// TIA Portal V20 export
// export: Created 2026-10-20T12:39:45.8971226Z, ExportSetting WithDefaults, DisplayName Totally Integrated Automation Portal, DisplayVersion V20 Update 6, DisplayName TIA Portal Openness, DisplayVersion V20 Update 6, DisplayName TIA Portal Version Control Interface, DisplayVersion V20 Update 6, DisplayName SINAMICS Startdrive Advanced, DisplayVersion V20 SP1, DisplayName SINAMICS Startdrive G130, G150, S120, S150, SINAMICS MV, G220, S200, S210, DisplayVersion V20 SP1, DisplayName SINAMICS Startdrive G110M, G120, G120C, G120D, G120P, G115D, DisplayVersion V20 SP1, DisplayName STEP 7 Professional, DisplayVersion V20 Update 6, DisplayName STEP 7 Safety, DisplayVersion V20 Update 2, DisplayName WinCC Basic/Comfort/Advanced, DisplayVersion V20 Update 6, DisplayName WinCC Unified, DisplayVersion V20 Update 6
FUNCTION_BLOCK "Main_Safety_RTG1"   // FB123, F_FBD
{ S7_Optimized_Access := 'TRUE' }
VERSION : 0.1
// stored: AutoNumber false, IsIECCheckEnabled false, UDAEnableTagReadback false
   VAR
      Safety_OK : Bool;
      ACK : Bool;
   END_VAR
   VAR_TEMP
      HMI_1_Estop_Pressed_1 : Bool;
      HMI_1_Estop_Pressed_2 : Bool;
      HMI_1_Estop_Pressed_3 : Bool;
      HMI_1_Estop_Pressed_4 : Bool;
      HMI_1_Estop_Pressed_5 : Bool;
      HMI_2_Estop_Pressed_1 : Bool;
      HMI_2_Estop_Pressed_2 : Bool;
      HMI_2_Estop_Pressed_3 : Bool;
      HMI_2_Estop_Pressed_4 : Bool;
      HMI_2_Estop_Pressed_5 : Bool;
      HMI_1_Reset_Comiss_1 : Bool;
      HMI_1_Reset_Comiss_2 : Bool;
      HMI_1_Reset_Comiss_3 : Bool;
      HMI_1_Reset_Comiss_4 : Bool;
      HMI_1_Reset_Comiss_5 : Bool;
      HMI_2_Reset_Comiss_1 : Bool;
      HMI_2_Reset_Comiss_2 : Bool;
      HMI_2_Reset_Comiss_3 : Bool;
      HMI_2_Reset_Comiss_4 : Bool;
      HMI_2_Reset_Comiss_5 : Bool;
   END_VAR
BEGIN

REGION Network 1: MAIN PANEL
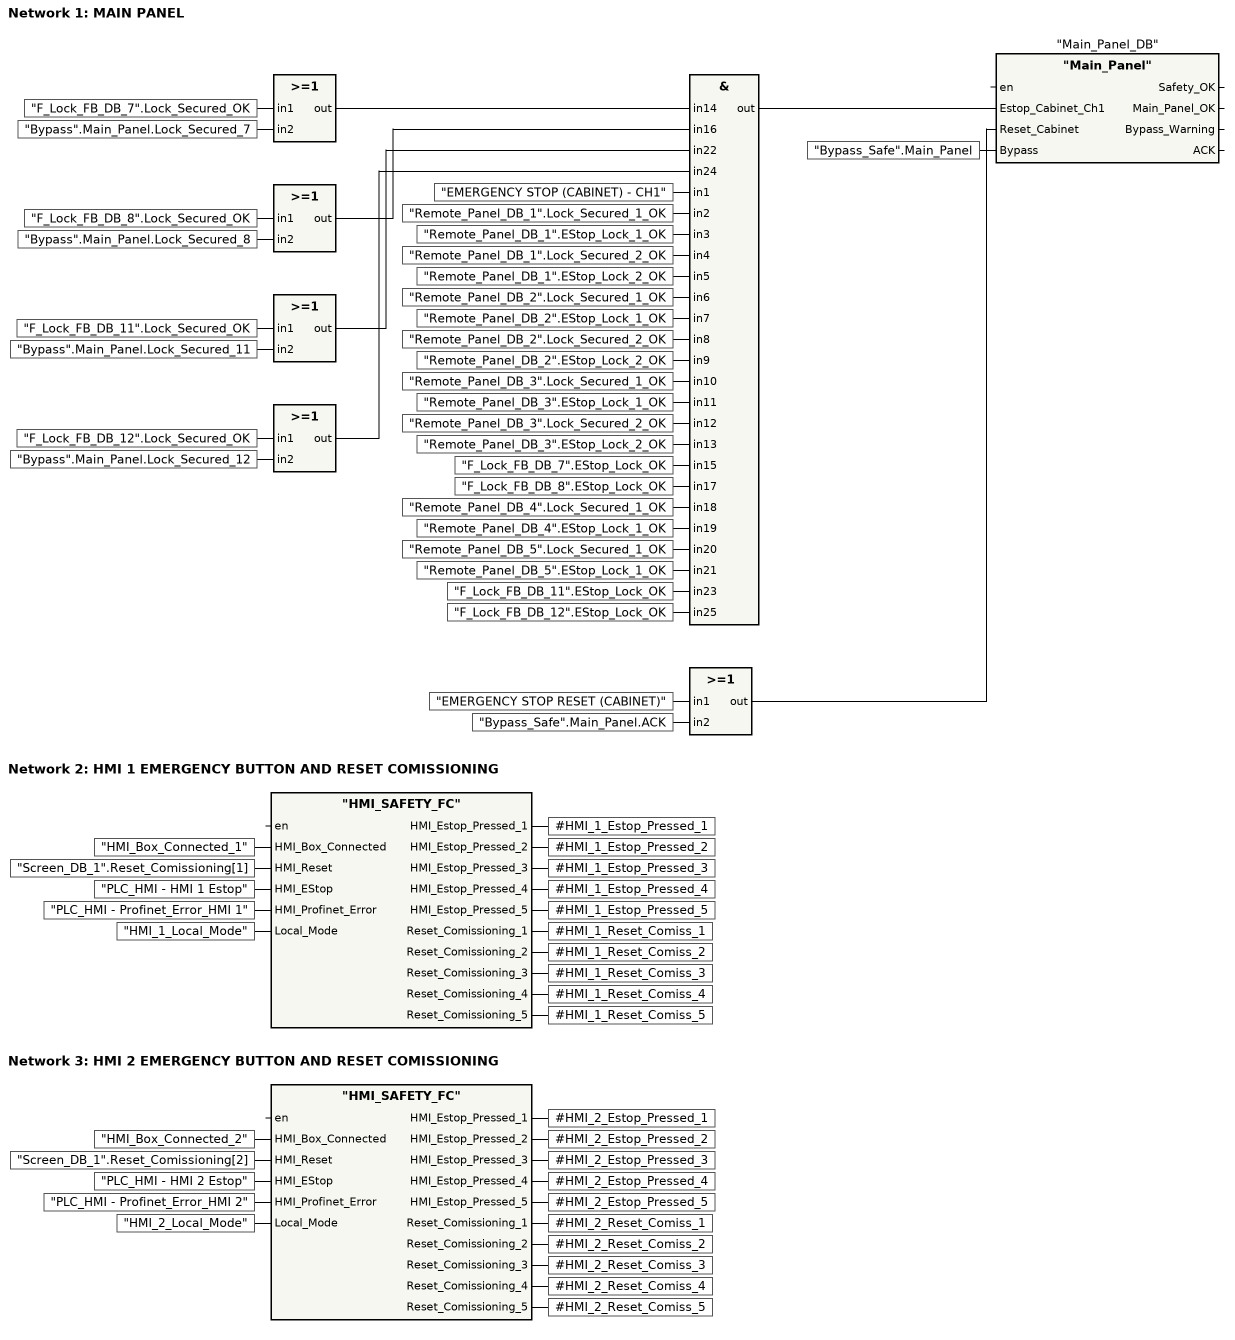
   "Main_Panel_DB"(Estop_Cabinet_Ch1 := ("F_Lock_FB_DB_7".Lock_Secured_OK OR "Bypass".Main_Panel.Lock_Secured_7) AND ("F_Lock_FB_DB_8".Lock_Secured_OK OR "Bypass".Main_Panel.Lock_Secured_8) AND ("F_Lock_FB_DB_11".Lock_Secured_OK OR "Bypass".Main_Panel.Lock_Secured_11) AND ("F_Lock_FB_DB_12".Lock_Secured_OK OR "Bypass".Main_Panel.Lock_Secured_12) AND "EMERGENCY STOP (CABINET) - CH1" AND "Remote_Panel_DB_1".Lock_Secured_1_OK AND "Remote_Panel_DB_1".EStop_Lock_1_OK AND "Remote_Panel_DB_1".Lock_Secured_2_OK AND "Remote_Panel_DB_1".EStop_Lock_2_OK AND "Remote_Panel_DB_2".Lock_Secured_1_OK AND "Remote_Panel_DB_2".EStop_Lock_1_OK AND "Remote_Panel_DB_2".Lock_Secured_2_OK AND "Remote_Panel_DB_2".EStop_Lock_2_OK AND "Remote_Panel_DB_3".Lock_Secured_1_OK AND "Remote_Panel_DB_3".EStop_Lock_1_OK AND "Remote_Panel_DB_3".Lock_Secured_2_OK AND "Remote_Panel_DB_3".EStop_Lock_2_OK AND "F_Lock_FB_DB_7".EStop_Lock_OK AND "F_Lock_FB_DB_8".EStop_Lock_OK AND "Remote_Panel_DB_4".Lock_Secured_1_OK AND "Remote_Panel_DB_4".EStop_Lock_1_OK AND "Remote_Panel_DB_5".Lock_Secured_1_OK AND "Remote_Panel_DB_5".EStop_Lock_1_OK AND "F_Lock_FB_DB_11".EStop_Lock_OK AND "F_Lock_FB_DB_12".EStop_Lock_OK,   // "Main_Panel"
                   Reset_Cabinet := "EMERGENCY STOP RESET (CABINET)" OR "Bypass_Safe".Main_Panel.ACK,
                   Bypass := "Bypass_Safe".Main_Panel);
END_REGION

REGION Network 2: HMI 1 EMERGENCY BUTTON AND RESET COMISSIONING
   "HMI_SAFETY_FC"(HMI_Box_Connected := "HMI_Box_Connected_1",
                   HMI_Reset := "Screen_DB_1".Reset_Comissioning[1],
                   HMI_EStop := "PLC_HMI - HMI 1 Estop",
                   HMI_Profinet_Error := "PLC_HMI - Profinet_Error_HMI 1",
                   Local_Mode := "HMI_1_Local_Mode",
                   HMI_Estop_Pressed_1 => #HMI_1_Estop_Pressed_1,
                   HMI_Estop_Pressed_2 => #HMI_1_Estop_Pressed_2,
                   HMI_Estop_Pressed_3 => #HMI_1_Estop_Pressed_3,
                   HMI_Estop_Pressed_4 => #HMI_1_Estop_Pressed_4,
                   HMI_Estop_Pressed_5 => #HMI_1_Estop_Pressed_5,
                   Reset_Comissioning_1 => #HMI_1_Reset_Comiss_1,
                   Reset_Comissioning_2 => #HMI_1_Reset_Comiss_2,
                   Reset_Comissioning_3 => #HMI_1_Reset_Comiss_3,
                   Reset_Comissioning_4 => #HMI_1_Reset_Comiss_4,
                   Reset_Comissioning_5 => #HMI_1_Reset_Comiss_5);
END_REGION

REGION Network 3: HMI 2 EMERGENCY BUTTON AND RESET COMISSIONING
   "HMI_SAFETY_FC"(HMI_Box_Connected := "HMI_Box_Connected_2",
                   HMI_Reset := "Screen_DB_1".Reset_Comissioning[2],
                   HMI_EStop := "PLC_HMI - HMI 2 Estop",
                   HMI_Profinet_Error := "PLC_HMI - Profinet_Error_HMI 2",
                   Local_Mode := "HMI_2_Local_Mode",
                   HMI_Estop_Pressed_1 => #HMI_2_Estop_Pressed_1,
                   HMI_Estop_Pressed_2 => #HMI_2_Estop_Pressed_2,
                   HMI_Estop_Pressed_3 => #HMI_2_Estop_Pressed_3,
                   HMI_Estop_Pressed_4 => #HMI_2_Estop_Pressed_4,
                   HMI_Estop_Pressed_5 => #HMI_2_Estop_Pressed_5,
                   Reset_Comissioning_1 => #HMI_2_Reset_Comiss_1,
                   Reset_Comissioning_2 => #HMI_2_Reset_Comiss_2,
                   Reset_Comissioning_3 => #HMI_2_Reset_Comiss_3,
                   Reset_Comissioning_4 => #HMI_2_Reset_Comiss_4,
                   Reset_Comissioning_5 => #HMI_2_Reset_Comiss_5);
END_REGION

REGION Network 4: Remote Panel 1
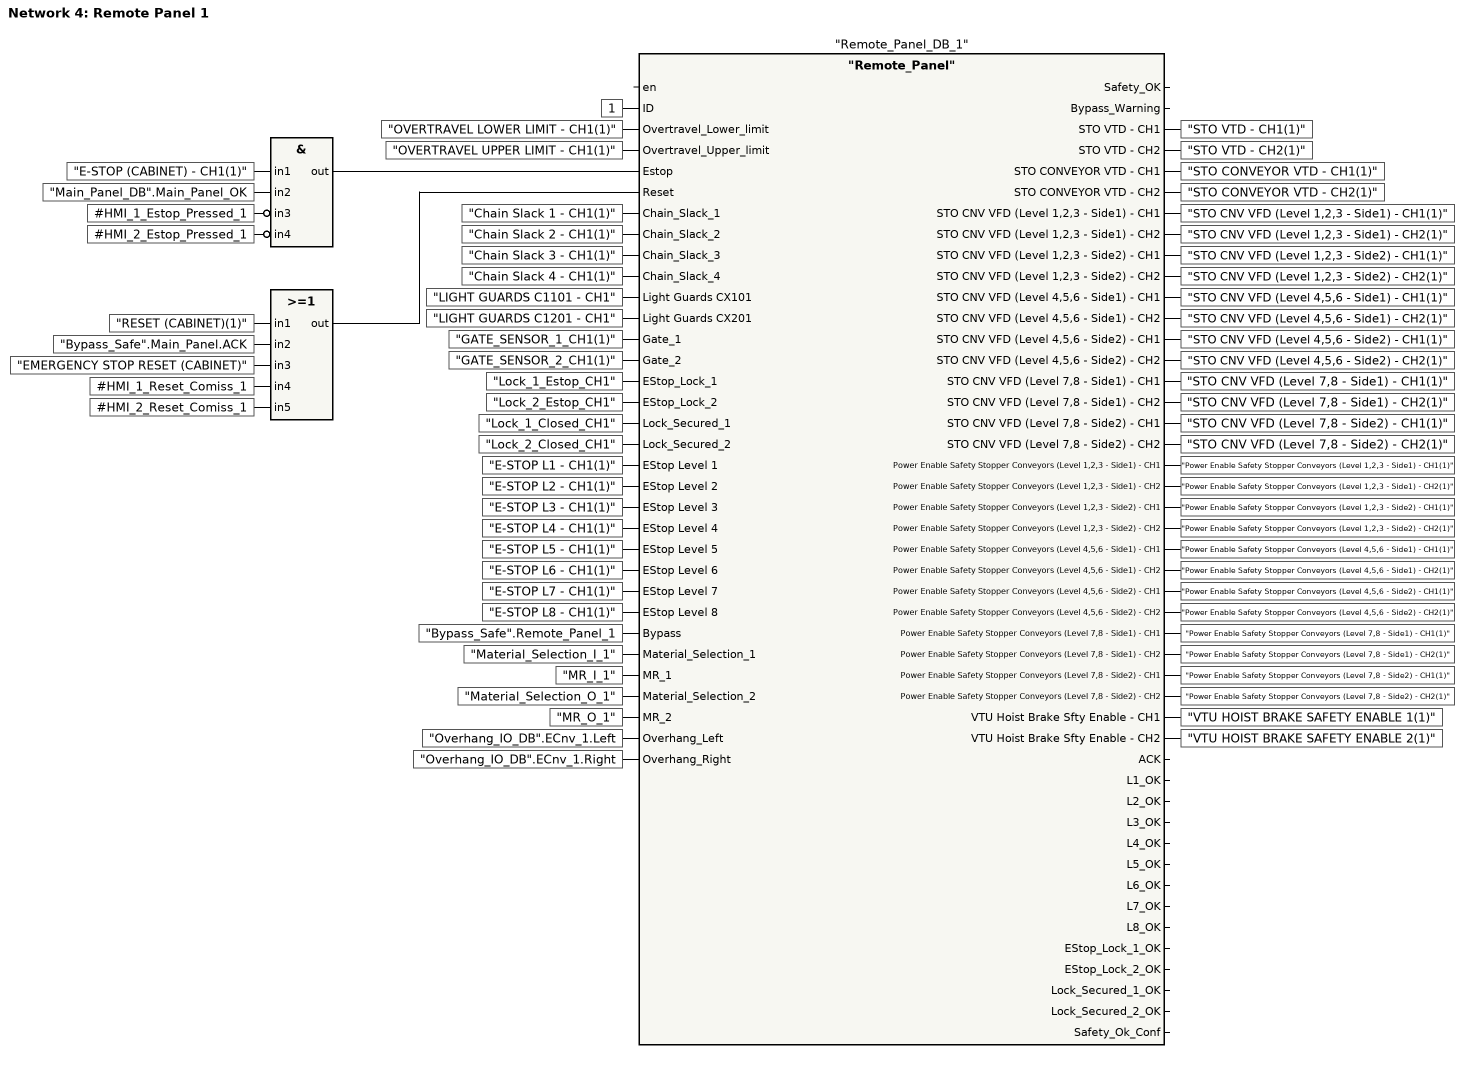
   "Remote_Panel_DB_1"(ID := 1,   // "Remote_Panel"
                       Overtravel_Lower_limit := "OVERTRAVEL LOWER LIMIT - CH1(1)",
                       Overtravel_Upper_limit := "OVERTRAVEL UPPER LIMIT - CH1(1)",
                       Estop := "E-STOP (CABINET) - CH1(1)" AND "Main_Panel_DB".Main_Panel_OK AND NOT #HMI_1_Estop_Pressed_1 AND NOT #HMI_2_Estop_Pressed_1,
                       Reset := "RESET (CABINET)(1)" OR "Bypass_Safe".Main_Panel.ACK OR "EMERGENCY STOP RESET (CABINET)" OR #HMI_1_Reset_Comiss_1 OR #HMI_2_Reset_Comiss_1,
                       Chain_Slack_1 := "Chain Slack 1 - CH1(1)",
                       Chain_Slack_2 := "Chain Slack 2 - CH1(1)",
                       Chain_Slack_3 := "Chain Slack 3 - CH1(1)",
                       Chain_Slack_4 := "Chain Slack 4 - CH1(1)",
                       "Light Guards CX101" := "LIGHT GUARDS C1101 - CH1",
                       "Light Guards CX201" := "LIGHT GUARDS C1201 - CH1",
                       Gate_1 := "GATE_SENSOR_1_CH1(1)",
                       Gate_2 := "GATE_SENSOR_2_CH1(1)",
                       EStop_Lock_1 := "Lock_1_Estop_CH1",
                       EStop_Lock_2 := "Lock_2_Estop_CH1",
                       Lock_Secured_1 := "Lock_1_Closed_CH1",
                       Lock_Secured_2 := "Lock_2_Closed_CH1",
                       "EStop Level 1" := "E-STOP L1 - CH1(1)",
                       "EStop Level 2" := "E-STOP L2 - CH1(1)",
                       "EStop Level 3" := "E-STOP L3 - CH1(1)",
                       "EStop Level 4" := "E-STOP L4 - CH1(1)",
                       "EStop Level 5" := "E-STOP L5 - CH1(1)",
                       "EStop Level 6" := "E-STOP L6 - CH1(1)",
                       "EStop Level 7" := "E-STOP L7 - CH1(1)",
                       "EStop Level 8" := "E-STOP L8 - CH1(1)",
                       Bypass := "Bypass_Safe".Remote_Panel_1,
                       Material_Selection_1 := "Material_Selection_I_1",
                       MR_1 := "MR_I_1",
                       Material_Selection_2 := "Material_Selection_O_1",
                       MR_2 := "MR_O_1",
                       Overhang_Left := "Overhang_IO_DB".ECnv_1.Left,
                       Overhang_Right := "Overhang_IO_DB".ECnv_1.Right,
                       "STO VTD - CH1" => "STO VTD - CH1(1)",
                       "STO VTD - CH2" => "STO VTD - CH2(1)",
                       "STO CONVEYOR VTD - CH1" => "STO CONVEYOR VTD - CH1(1)",
                       "STO CONVEYOR VTD - CH2" => "STO CONVEYOR VTD - CH2(1)",
                       "STO CNV VFD (Level 1,2,3 - Side1) - CH1" => "STO CNV VFD (Level 1,2,3 - Side1) - CH1(1)",
                       "STO CNV VFD (Level 1,2,3 - Side1) - CH2" => "STO CNV VFD (Level 1,2,3 - Side1) - CH2(1)",
                       "STO CNV VFD (Level 1,2,3 - Side2) - CH1" => "STO CNV VFD (Level 1,2,3 - Side2) - CH1(1)",
                       "STO CNV VFD (Level 1,2,3 - Side2) - CH2" => "STO CNV VFD (Level 1,2,3 - Side2) - CH2(1)",
                       "STO CNV VFD (Level 4,5,6 - Side1) - CH1" => "STO CNV VFD (Level 4,5,6 - Side1) - CH1(1)",
                       "STO CNV VFD (Level 4,5,6 - Side1) - CH2" => "STO CNV VFD (Level 4,5,6 - Side1) - CH2(1)",
                       "STO CNV VFD (Level 4,5,6 - Side2) - CH1" => "STO CNV VFD (Level 4,5,6 - Side2) - CH1(1)",
                       "STO CNV VFD (Level 4,5,6 - Side2) - CH2" => "STO CNV VFD (Level 4,5,6 - Side2) - CH2(1)",
                       "STO CNV VFD (Level 7,8 - Side1) - CH1" => "STO CNV VFD (Level 7,8 - Side1) - CH1(1)",
                       "STO CNV VFD (Level 7,8 - Side1) - CH2" => "STO CNV VFD (Level 7,8 - Side1) - CH2(1)",
                       "STO CNV VFD (Level 7,8 - Side2) - CH1" => "STO CNV VFD (Level 7,8 - Side2) - CH1(1)",
                       "STO CNV VFD (Level 7,8 - Side2) - CH2" => "STO CNV VFD (Level 7,8 - Side2) - CH2(1)",
                       "Power Enable Safety Stopper Conveyors (Level 1,2,3 - Side1) - CH1" => "Power Enable Safety Stopper Conveyors (Level 1,2,3 - Side1) - CH1(1)",
                       "Power Enable Safety Stopper Conveyors (Level 1,2,3 - Side1) - CH2" => "Power Enable Safety Stopper Conveyors (Level 1,2,3 - Side1) - CH2(1)",
                       "Power Enable Safety Stopper Conveyors (Level 1,2,3 - Side2) - CH1" => "Power Enable Safety Stopper Conveyors (Level 1,2,3 - Side2) - CH1(1)",
                       "Power Enable Safety Stopper Conveyors (Level 1,2,3 - Side2) - CH2" => "Power Enable Safety Stopper Conveyors (Level 1,2,3 - Side2) - CH2(1)",
                       "Power Enable Safety Stopper Conveyors (Level 4,5,6 - Side1) - CH1" => "Power Enable Safety Stopper Conveyors (Level 4,5,6 - Side1) - CH1(1)",
                       "Power Enable Safety Stopper Conveyors (Level 4,5,6 - Side1) - CH2" => "Power Enable Safety Stopper Conveyors (Level 4,5,6 - Side1) - CH2(1)",
                       "Power Enable Safety Stopper Conveyors (Level 4,5,6 - Side2) - CH1" => "Power Enable Safety Stopper Conveyors (Level 4,5,6 - Side2) - CH1(1)",
                       "Power Enable Safety Stopper Conveyors (Level 4,5,6 - Side2) - CH2" => "Power Enable Safety Stopper Conveyors (Level 4,5,6 - Side2) - CH2(1)",
                       "Power Enable Safety Stopper Conveyors (Level 7,8 - Side1) - CH1" => "Power Enable Safety Stopper Conveyors (Level 7,8 - Side1) - CH1(1)",
                       "Power Enable Safety Stopper Conveyors (Level 7,8 - Side1) - CH2" => "Power Enable Safety Stopper Conveyors (Level 7,8 - Side1) - CH2(1)",
                       "Power Enable Safety Stopper Conveyors (Level 7,8 - Side2) - CH1" => "Power Enable Safety Stopper Conveyors (Level 7,8 - Side2) - CH1(1)",
                       "Power Enable Safety Stopper Conveyors (Level 7,8 - Side2) - CH2" => "Power Enable Safety Stopper Conveyors (Level 7,8 - Side2) - CH2(1)",
                       "VTU Hoist Brake Sfty Enable - CH1" => "VTU HOIST BRAKE SAFETY ENABLE 1(1)",
                       "VTU Hoist Brake Sfty Enable - CH2" => "VTU HOIST BRAKE SAFETY ENABLE 2(1)");
END_REGION

REGION Network 5: Remote Panel 2
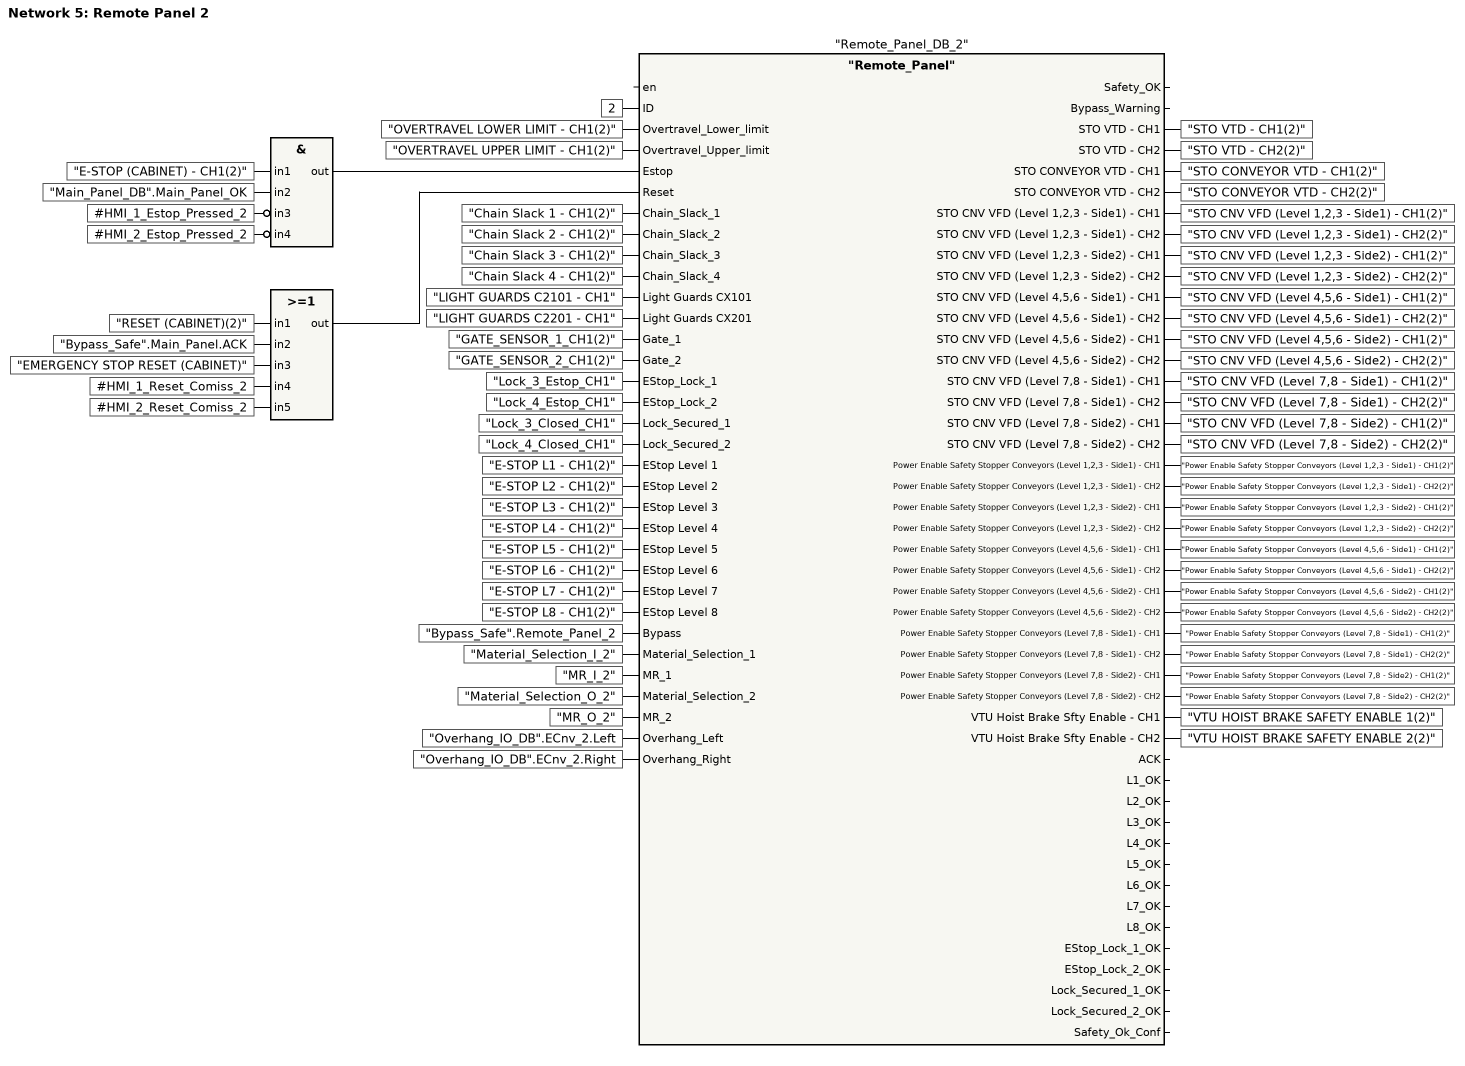
   "Remote_Panel_DB_2"(ID := 2,   // "Remote_Panel"
                       Overtravel_Lower_limit := "OVERTRAVEL LOWER LIMIT - CH1(2)",
                       Overtravel_Upper_limit := "OVERTRAVEL UPPER LIMIT - CH1(2)",
                       Estop := "E-STOP (CABINET) - CH1(2)" AND "Main_Panel_DB".Main_Panel_OK AND NOT #HMI_1_Estop_Pressed_2 AND NOT #HMI_2_Estop_Pressed_2,
                       Reset := "RESET (CABINET)(2)" OR "Bypass_Safe".Main_Panel.ACK OR "EMERGENCY STOP RESET (CABINET)" OR #HMI_1_Reset_Comiss_2 OR #HMI_2_Reset_Comiss_2,
                       Chain_Slack_1 := "Chain Slack 1 - CH1(2)",
                       Chain_Slack_2 := "Chain Slack 2 - CH1(2)",
                       Chain_Slack_3 := "Chain Slack 3 - CH1(2)",
                       Chain_Slack_4 := "Chain Slack 4 - CH1(2)",
                       "Light Guards CX101" := "LIGHT GUARDS C2101 - CH1",
                       "Light Guards CX201" := "LIGHT GUARDS C2201 - CH1",
                       Gate_1 := "GATE_SENSOR_1_CH1(2)",
                       Gate_2 := "GATE_SENSOR_2_CH1(2)",
                       EStop_Lock_1 := "Lock_3_Estop_CH1",
                       EStop_Lock_2 := "Lock_4_Estop_CH1",
                       Lock_Secured_1 := "Lock_3_Closed_CH1",
                       Lock_Secured_2 := "Lock_4_Closed_CH1",
                       "EStop Level 1" := "E-STOP L1 - CH1(2)",
                       "EStop Level 2" := "E-STOP L2 - CH1(2)",
                       "EStop Level 3" := "E-STOP L3 - CH1(2)",
                       "EStop Level 4" := "E-STOP L4 - CH1(2)",
                       "EStop Level 5" := "E-STOP L5 - CH1(2)",
                       "EStop Level 6" := "E-STOP L6 - CH1(2)",
                       "EStop Level 7" := "E-STOP L7 - CH1(2)",
                       "EStop Level 8" := "E-STOP L8 - CH1(2)",
                       Bypass := "Bypass_Safe".Remote_Panel_2,
                       Material_Selection_1 := "Material_Selection_I_2",
                       MR_1 := "MR_I_2",
                       Material_Selection_2 := "Material_Selection_O_2",
                       MR_2 := "MR_O_2",
                       Overhang_Left := "Overhang_IO_DB".ECnv_2.Left,
                       Overhang_Right := "Overhang_IO_DB".ECnv_2.Right,
                       "STO VTD - CH1" => "STO VTD - CH1(2)",
                       "STO VTD - CH2" => "STO VTD - CH2(2)",
                       "STO CONVEYOR VTD - CH1" => "STO CONVEYOR VTD - CH1(2)",
                       "STO CONVEYOR VTD - CH2" => "STO CONVEYOR VTD - CH2(2)",
                       "STO CNV VFD (Level 1,2,3 - Side1) - CH1" => "STO CNV VFD (Level 1,2,3 - Side1) - CH1(2)",
                       "STO CNV VFD (Level 1,2,3 - Side1) - CH2" => "STO CNV VFD (Level 1,2,3 - Side1) - CH2(2)",
                       "STO CNV VFD (Level 1,2,3 - Side2) - CH1" => "STO CNV VFD (Level 1,2,3 - Side2) - CH1(2)",
                       "STO CNV VFD (Level 1,2,3 - Side2) - CH2" => "STO CNV VFD (Level 1,2,3 - Side2) - CH2(2)",
                       "STO CNV VFD (Level 4,5,6 - Side1) - CH1" => "STO CNV VFD (Level 4,5,6 - Side1) - CH1(2)",
                       "STO CNV VFD (Level 4,5,6 - Side1) - CH2" => "STO CNV VFD (Level 4,5,6 - Side1) - CH2(2)",
                       "STO CNV VFD (Level 4,5,6 - Side2) - CH1" => "STO CNV VFD (Level 4,5,6 - Side2) - CH1(2)",
                       "STO CNV VFD (Level 4,5,6 - Side2) - CH2" => "STO CNV VFD (Level 4,5,6 - Side2) - CH2(2)",
                       "STO CNV VFD (Level 7,8 - Side1) - CH1" => "STO CNV VFD (Level 7,8 - Side1) - CH1(2)",
                       "STO CNV VFD (Level 7,8 - Side1) - CH2" => "STO CNV VFD (Level 7,8 - Side1) - CH2(2)",
                       "STO CNV VFD (Level 7,8 - Side2) - CH1" => "STO CNV VFD (Level 7,8 - Side2) - CH1(2)",
                       "STO CNV VFD (Level 7,8 - Side2) - CH2" => "STO CNV VFD (Level 7,8 - Side2) - CH2(2)",
                       "Power Enable Safety Stopper Conveyors (Level 1,2,3 - Side1) - CH1" => "Power Enable Safety Stopper Conveyors (Level 1,2,3 - Side1) - CH1(2)",
                       "Power Enable Safety Stopper Conveyors (Level 1,2,3 - Side1) - CH2" => "Power Enable Safety Stopper Conveyors (Level 1,2,3 - Side1) - CH2(2)",
                       "Power Enable Safety Stopper Conveyors (Level 1,2,3 - Side2) - CH1" => "Power Enable Safety Stopper Conveyors (Level 1,2,3 - Side2) - CH1(2)",
                       "Power Enable Safety Stopper Conveyors (Level 1,2,3 - Side2) - CH2" => "Power Enable Safety Stopper Conveyors (Level 1,2,3 - Side2) - CH2(2)",
                       "Power Enable Safety Stopper Conveyors (Level 4,5,6 - Side1) - CH1" => "Power Enable Safety Stopper Conveyors (Level 4,5,6 - Side1) - CH1(2)",
                       "Power Enable Safety Stopper Conveyors (Level 4,5,6 - Side1) - CH2" => "Power Enable Safety Stopper Conveyors (Level 4,5,6 - Side1) - CH2(2)",
                       "Power Enable Safety Stopper Conveyors (Level 4,5,6 - Side2) - CH1" => "Power Enable Safety Stopper Conveyors (Level 4,5,6 - Side2) - CH1(2)",
                       "Power Enable Safety Stopper Conveyors (Level 4,5,6 - Side2) - CH2" => "Power Enable Safety Stopper Conveyors (Level 4,5,6 - Side2) - CH2(2)",
                       "Power Enable Safety Stopper Conveyors (Level 7,8 - Side1) - CH1" => "Power Enable Safety Stopper Conveyors (Level 7,8 - Side1) - CH1(2)",
                       "Power Enable Safety Stopper Conveyors (Level 7,8 - Side1) - CH2" => "Power Enable Safety Stopper Conveyors (Level 7,8 - Side1) - CH2(2)",
                       "Power Enable Safety Stopper Conveyors (Level 7,8 - Side2) - CH1" => "Power Enable Safety Stopper Conveyors (Level 7,8 - Side2) - CH1(2)",
                       "Power Enable Safety Stopper Conveyors (Level 7,8 - Side2) - CH2" => "Power Enable Safety Stopper Conveyors (Level 7,8 - Side2) - CH2(2)",
                       "VTU Hoist Brake Sfty Enable - CH1" => "VTU HOIST BRAKE SAFETY ENABLE 1(2)",
                       "VTU Hoist Brake Sfty Enable - CH2" => "VTU HOIST BRAKE SAFETY ENABLE 2(2)");
END_REGION

REGION Network 6: Remote Panel 3
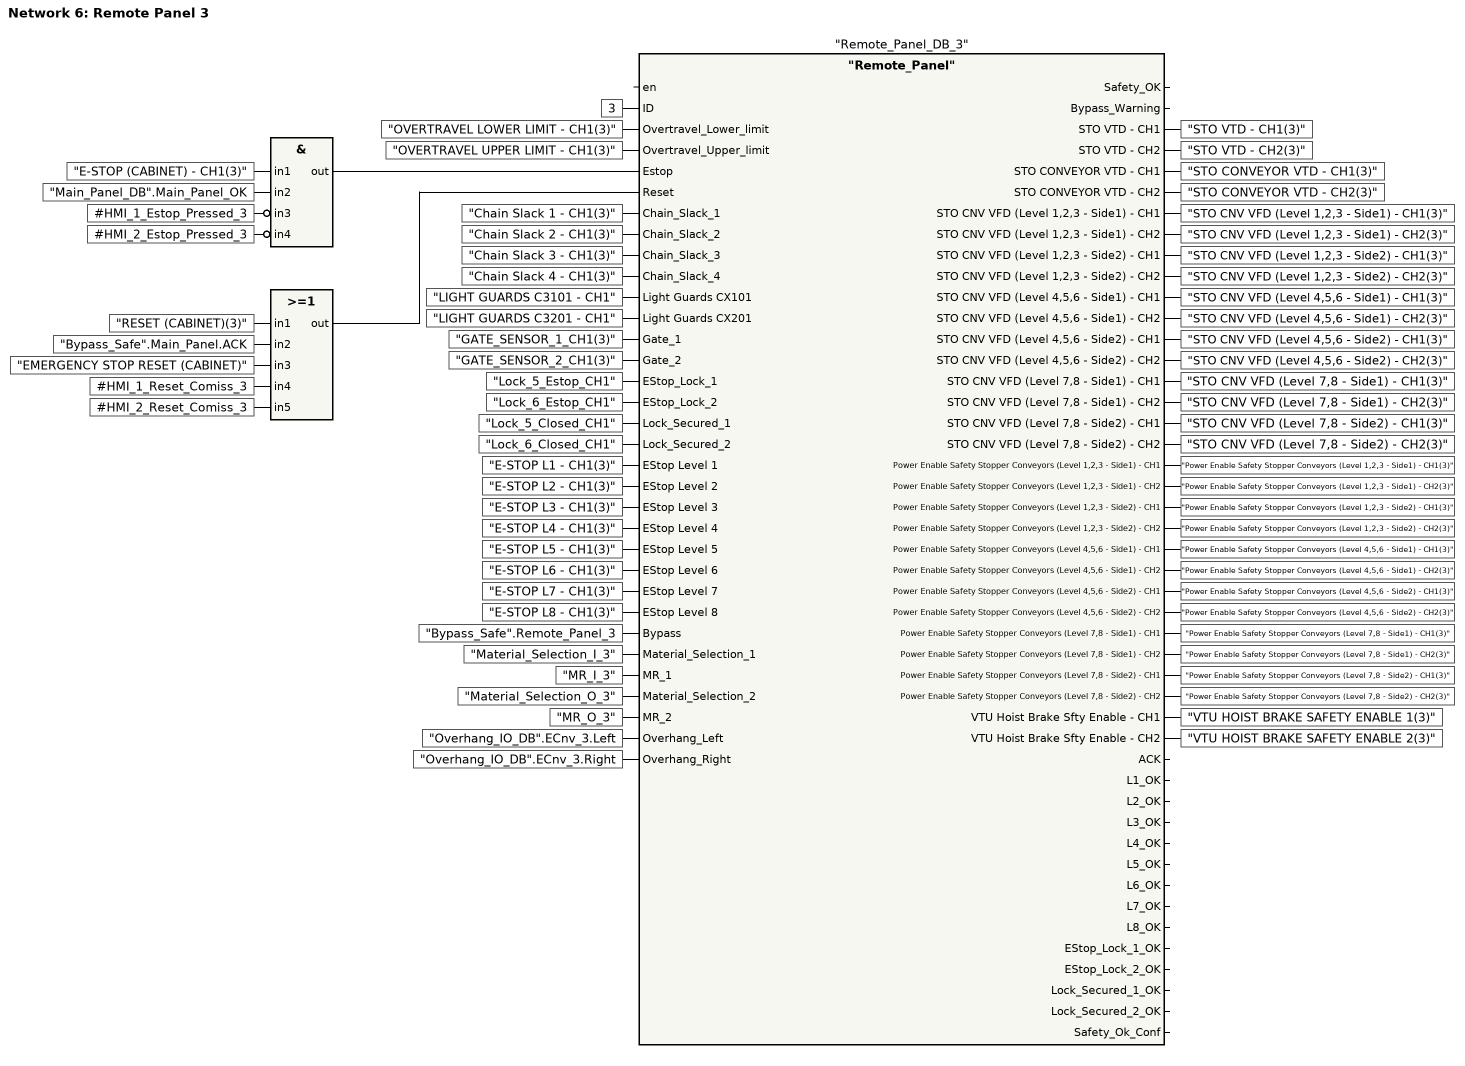
   "Remote_Panel_DB_3"(ID := 3,   // "Remote_Panel"
                       Overtravel_Lower_limit := "OVERTRAVEL LOWER LIMIT - CH1(3)",
                       Overtravel_Upper_limit := "OVERTRAVEL UPPER LIMIT - CH1(3)",
                       Estop := "E-STOP (CABINET) - CH1(3)" AND "Main_Panel_DB".Main_Panel_OK AND NOT #HMI_1_Estop_Pressed_3 AND NOT #HMI_2_Estop_Pressed_3,
                       Reset := "RESET (CABINET)(3)" OR "Bypass_Safe".Main_Panel.ACK OR "EMERGENCY STOP RESET (CABINET)" OR #HMI_1_Reset_Comiss_3 OR #HMI_2_Reset_Comiss_3,
                       Chain_Slack_1 := "Chain Slack 1 - CH1(3)",
                       Chain_Slack_2 := "Chain Slack 2 - CH1(3)",
                       Chain_Slack_3 := "Chain Slack 3 - CH1(3)",
                       Chain_Slack_4 := "Chain Slack 4 - CH1(3)",
                       "Light Guards CX101" := "LIGHT GUARDS C3101 - CH1",
                       "Light Guards CX201" := "LIGHT GUARDS C3201 - CH1",
                       Gate_1 := "GATE_SENSOR_1_CH1(3)",
                       Gate_2 := "GATE_SENSOR_2_CH1(3)",
                       EStop_Lock_1 := "Lock_5_Estop_CH1",
                       EStop_Lock_2 := "Lock_6_Estop_CH1",
                       Lock_Secured_1 := "Lock_5_Closed_CH1",
                       Lock_Secured_2 := "Lock_6_Closed_CH1",
                       "EStop Level 1" := "E-STOP L1 - CH1(3)",
                       "EStop Level 2" := "E-STOP L2 - CH1(3)",
                       "EStop Level 3" := "E-STOP L3 - CH1(3)",
                       "EStop Level 4" := "E-STOP L4 - CH1(3)",
                       "EStop Level 5" := "E-STOP L5 - CH1(3)",
                       "EStop Level 6" := "E-STOP L6 - CH1(3)",
                       "EStop Level 7" := "E-STOP L7 - CH1(3)",
                       "EStop Level 8" := "E-STOP L8 - CH1(3)",
                       Bypass := "Bypass_Safe".Remote_Panel_3,
                       Material_Selection_1 := "Material_Selection_I_3",
                       MR_1 := "MR_I_3",
                       Material_Selection_2 := "Material_Selection_O_3",
                       MR_2 := "MR_O_3",
                       Overhang_Left := "Overhang_IO_DB".ECnv_3.Left,
                       Overhang_Right := "Overhang_IO_DB".ECnv_3.Right,
                       "STO VTD - CH1" => "STO VTD - CH1(3)",
                       "STO VTD - CH2" => "STO VTD - CH2(3)",
                       "STO CONVEYOR VTD - CH1" => "STO CONVEYOR VTD - CH1(3)",
                       "STO CONVEYOR VTD - CH2" => "STO CONVEYOR VTD - CH2(3)",
                       "STO CNV VFD (Level 1,2,3 - Side1) - CH1" => "STO CNV VFD (Level 1,2,3 - Side1) - CH1(3)",
                       "STO CNV VFD (Level 1,2,3 - Side1) - CH2" => "STO CNV VFD (Level 1,2,3 - Side1) - CH2(3)",
                       "STO CNV VFD (Level 1,2,3 - Side2) - CH1" => "STO CNV VFD (Level 1,2,3 - Side2) - CH1(3)",
                       "STO CNV VFD (Level 1,2,3 - Side2) - CH2" => "STO CNV VFD (Level 1,2,3 - Side2) - CH2(3)",
                       "STO CNV VFD (Level 4,5,6 - Side1) - CH1" => "STO CNV VFD (Level 4,5,6 - Side1) - CH1(3)",
                       "STO CNV VFD (Level 4,5,6 - Side1) - CH2" => "STO CNV VFD (Level 4,5,6 - Side1) - CH2(3)",
                       "STO CNV VFD (Level 4,5,6 - Side2) - CH1" => "STO CNV VFD (Level 4,5,6 - Side2) - CH1(3)",
                       "STO CNV VFD (Level 4,5,6 - Side2) - CH2" => "STO CNV VFD (Level 4,5,6 - Side2) - CH2(3)",
                       "STO CNV VFD (Level 7,8 - Side1) - CH1" => "STO CNV VFD (Level 7,8 - Side1) - CH1(3)",
                       "STO CNV VFD (Level 7,8 - Side1) - CH2" => "STO CNV VFD (Level 7,8 - Side1) - CH2(3)",
                       "STO CNV VFD (Level 7,8 - Side2) - CH1" => "STO CNV VFD (Level 7,8 - Side2) - CH1(3)",
                       "STO CNV VFD (Level 7,8 - Side2) - CH2" => "STO CNV VFD (Level 7,8 - Side2) - CH2(3)",
                       "Power Enable Safety Stopper Conveyors (Level 1,2,3 - Side1) - CH1" => "Power Enable Safety Stopper Conveyors (Level 1,2,3 - Side1) - CH1(3)",
                       "Power Enable Safety Stopper Conveyors (Level 1,2,3 - Side1) - CH2" => "Power Enable Safety Stopper Conveyors (Level 1,2,3 - Side1) - CH2(3)",
                       "Power Enable Safety Stopper Conveyors (Level 1,2,3 - Side2) - CH1" => "Power Enable Safety Stopper Conveyors (Level 1,2,3 - Side2) - CH1(3)",
                       "Power Enable Safety Stopper Conveyors (Level 1,2,3 - Side2) - CH2" => "Power Enable Safety Stopper Conveyors (Level 1,2,3 - Side2) - CH2(3)",
                       "Power Enable Safety Stopper Conveyors (Level 4,5,6 - Side1) - CH1" => "Power Enable Safety Stopper Conveyors (Level 4,5,6 - Side1) - CH1(3)",
                       "Power Enable Safety Stopper Conveyors (Level 4,5,6 - Side1) - CH2" => "Power Enable Safety Stopper Conveyors (Level 4,5,6 - Side1) - CH2(3)",
                       "Power Enable Safety Stopper Conveyors (Level 4,5,6 - Side2) - CH1" => "Power Enable Safety Stopper Conveyors (Level 4,5,6 - Side2) - CH1(3)",
                       "Power Enable Safety Stopper Conveyors (Level 4,5,6 - Side2) - CH2" => "Power Enable Safety Stopper Conveyors (Level 4,5,6 - Side2) - CH2(3)",
                       "Power Enable Safety Stopper Conveyors (Level 7,8 - Side1) - CH1" => "Power Enable Safety Stopper Conveyors (Level 7,8 - Side1) - CH1(3)",
                       "Power Enable Safety Stopper Conveyors (Level 7,8 - Side1) - CH2" => "Power Enable Safety Stopper Conveyors (Level 7,8 - Side1) - CH2(3)",
                       "Power Enable Safety Stopper Conveyors (Level 7,8 - Side2) - CH1" => "Power Enable Safety Stopper Conveyors (Level 7,8 - Side2) - CH1(3)",
                       "Power Enable Safety Stopper Conveyors (Level 7,8 - Side2) - CH2" => "Power Enable Safety Stopper Conveyors (Level 7,8 - Side2) - CH2(3)",
                       "VTU Hoist Brake Sfty Enable - CH1" => "VTU HOIST BRAKE SAFETY ENABLE 1(3)",
                       "VTU Hoist Brake Sfty Enable - CH2" => "VTU HOIST BRAKE SAFETY ENABLE 2(3)");
END_REGION

REGION Network 7: Remote Panel 4
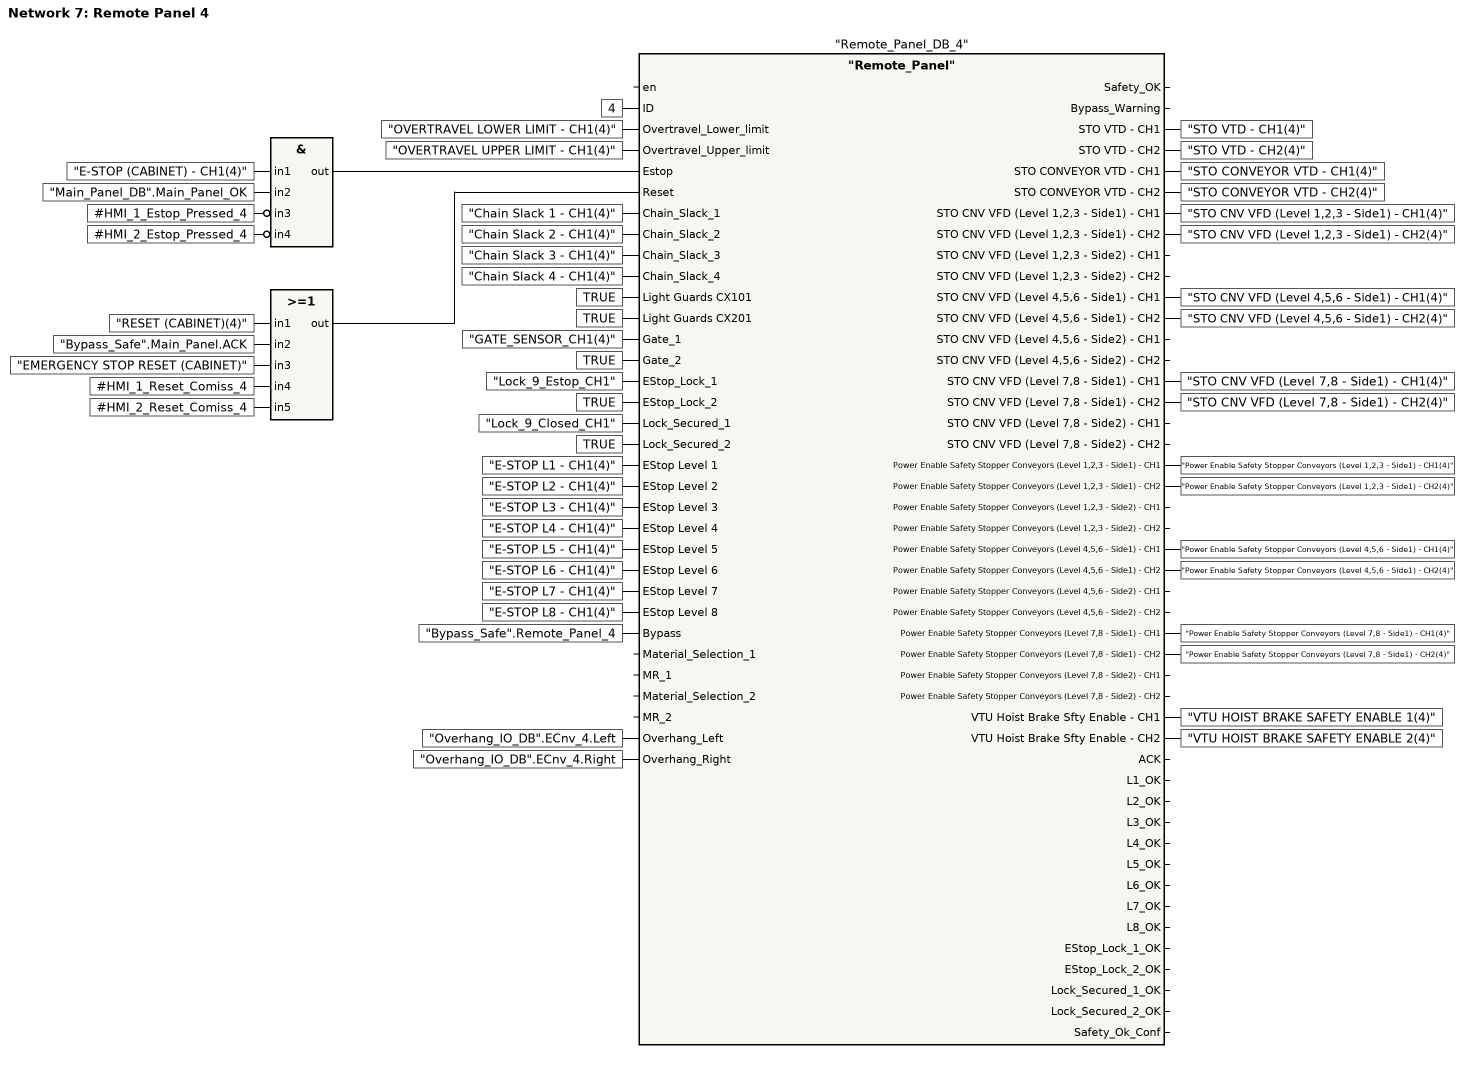
   "Remote_Panel_DB_4"(ID := 4,   // "Remote_Panel"
                       Overtravel_Lower_limit := "OVERTRAVEL LOWER LIMIT - CH1(4)",
                       Overtravel_Upper_limit := "OVERTRAVEL UPPER LIMIT - CH1(4)",
                       Estop := "E-STOP (CABINET) - CH1(4)" AND "Main_Panel_DB".Main_Panel_OK AND NOT #HMI_1_Estop_Pressed_4 AND NOT #HMI_2_Estop_Pressed_4,
                       Reset := "RESET (CABINET)(4)" OR "Bypass_Safe".Main_Panel.ACK OR "EMERGENCY STOP RESET (CABINET)" OR #HMI_1_Reset_Comiss_4 OR #HMI_2_Reset_Comiss_4,
                       Chain_Slack_1 := "Chain Slack 1 - CH1(4)",
                       Chain_Slack_2 := "Chain Slack 2 - CH1(4)",
                       Chain_Slack_3 := "Chain Slack 3 - CH1(4)",
                       Chain_Slack_4 := "Chain Slack 4 - CH1(4)",
                       "Light Guards CX101" := TRUE,
                       "Light Guards CX201" := TRUE,
                       Gate_1 := "GATE_SENSOR_CH1(4)",
                       Gate_2 := TRUE,
                       EStop_Lock_1 := "Lock_9_Estop_CH1",
                       EStop_Lock_2 := TRUE,
                       Lock_Secured_1 := "Lock_9_Closed_CH1",
                       Lock_Secured_2 := TRUE,
                       "EStop Level 1" := "E-STOP L1 - CH1(4)",
                       "EStop Level 2" := "E-STOP L2 - CH1(4)",
                       "EStop Level 3" := "E-STOP L3 - CH1(4)",
                       "EStop Level 4" := "E-STOP L4 - CH1(4)",
                       "EStop Level 5" := "E-STOP L5 - CH1(4)",
                       "EStop Level 6" := "E-STOP L6 - CH1(4)",
                       "EStop Level 7" := "E-STOP L7 - CH1(4)",
                       "EStop Level 8" := "E-STOP L8 - CH1(4)",
                       Bypass := "Bypass_Safe".Remote_Panel_4,
                       Overhang_Left := "Overhang_IO_DB".ECnv_4.Left,
                       Overhang_Right := "Overhang_IO_DB".ECnv_4.Right,
                       "STO VTD - CH1" => "STO VTD - CH1(4)",
                       "STO VTD - CH2" => "STO VTD - CH2(4)",
                       "STO CONVEYOR VTD - CH1" => "STO CONVEYOR VTD - CH1(4)",
                       "STO CONVEYOR VTD - CH2" => "STO CONVEYOR VTD - CH2(4)",
                       "STO CNV VFD (Level 1,2,3 - Side1) - CH1" => "STO CNV VFD (Level 1,2,3 - Side1) - CH1(4)",
                       "STO CNV VFD (Level 1,2,3 - Side1) - CH2" => "STO CNV VFD (Level 1,2,3 - Side1) - CH2(4)",
                       "STO CNV VFD (Level 4,5,6 - Side1) - CH1" => "STO CNV VFD (Level 4,5,6 - Side1) - CH1(4)",
                       "STO CNV VFD (Level 4,5,6 - Side1) - CH2" => "STO CNV VFD (Level 4,5,6 - Side1) - CH2(4)",
                       "STO CNV VFD (Level 7,8 - Side1) - CH1" => "STO CNV VFD (Level 7,8 - Side1) - CH1(4)",
                       "STO CNV VFD (Level 7,8 - Side1) - CH2" => "STO CNV VFD (Level 7,8 - Side1) - CH2(4)",
                       "Power Enable Safety Stopper Conveyors (Level 1,2,3 - Side1) - CH1" => "Power Enable Safety Stopper Conveyors (Level 1,2,3 - Side1) - CH1(4)",
                       "Power Enable Safety Stopper Conveyors (Level 1,2,3 - Side1) - CH2" => "Power Enable Safety Stopper Conveyors (Level 1,2,3 - Side1) - CH2(4)",
                       "Power Enable Safety Stopper Conveyors (Level 4,5,6 - Side1) - CH1" => "Power Enable Safety Stopper Conveyors (Level 4,5,6 - Side1) - CH1(4)",
                       "Power Enable Safety Stopper Conveyors (Level 4,5,6 - Side1) - CH2" => "Power Enable Safety Stopper Conveyors (Level 4,5,6 - Side1) - CH2(4)",
                       "Power Enable Safety Stopper Conveyors (Level 7,8 - Side1) - CH1" => "Power Enable Safety Stopper Conveyors (Level 7,8 - Side1) - CH1(4)",
                       "Power Enable Safety Stopper Conveyors (Level 7,8 - Side1) - CH2" => "Power Enable Safety Stopper Conveyors (Level 7,8 - Side1) - CH2(4)",
                       "VTU Hoist Brake Sfty Enable - CH1" => "VTU HOIST BRAKE SAFETY ENABLE 1(4)",
                       "VTU Hoist Brake Sfty Enable - CH2" => "VTU HOIST BRAKE SAFETY ENABLE 2(4)");
END_REGION

REGION Network 8: Remote Panel 5
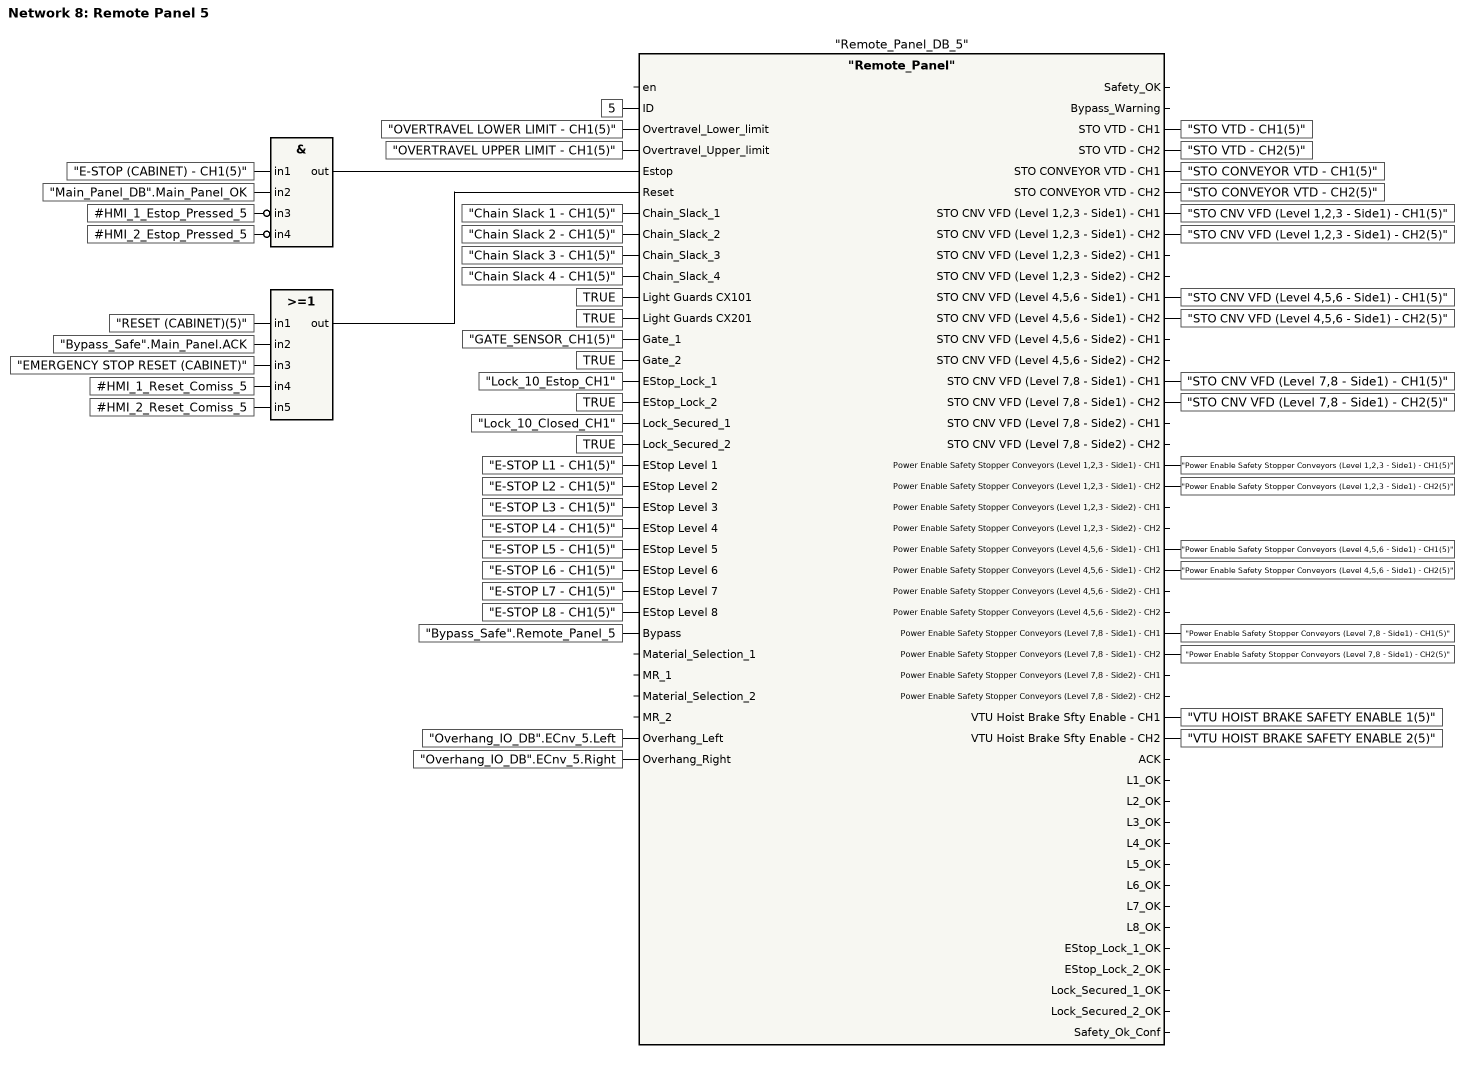
   "Remote_Panel_DB_5"(ID := 5,   // "Remote_Panel"
                       Overtravel_Lower_limit := "OVERTRAVEL LOWER LIMIT - CH1(5)",
                       Overtravel_Upper_limit := "OVERTRAVEL UPPER LIMIT - CH1(5)",
                       Estop := "E-STOP (CABINET) - CH1(5)" AND "Main_Panel_DB".Main_Panel_OK AND NOT #HMI_1_Estop_Pressed_5 AND NOT #HMI_2_Estop_Pressed_5,
                       Reset := "RESET (CABINET)(5)" OR "Bypass_Safe".Main_Panel.ACK OR "EMERGENCY STOP RESET (CABINET)" OR #HMI_1_Reset_Comiss_5 OR #HMI_2_Reset_Comiss_5,
                       Chain_Slack_1 := "Chain Slack 1 - CH1(5)",
                       Chain_Slack_2 := "Chain Slack 2 - CH1(5)",
                       Chain_Slack_3 := "Chain Slack 3 - CH1(5)",
                       Chain_Slack_4 := "Chain Slack 4 - CH1(5)",
                       "Light Guards CX101" := TRUE,
                       "Light Guards CX201" := TRUE,
                       Gate_1 := "GATE_SENSOR_CH1(5)",
                       Gate_2 := TRUE,
                       EStop_Lock_1 := "Lock_10_Estop_CH1",
                       EStop_Lock_2 := TRUE,
                       Lock_Secured_1 := "Lock_10_Closed_CH1",
                       Lock_Secured_2 := TRUE,
                       "EStop Level 1" := "E-STOP L1 - CH1(5)",
                       "EStop Level 2" := "E-STOP L2 - CH1(5)",
                       "EStop Level 3" := "E-STOP L3 - CH1(5)",
                       "EStop Level 4" := "E-STOP L4 - CH1(5)",
                       "EStop Level 5" := "E-STOP L5 - CH1(5)",
                       "EStop Level 6" := "E-STOP L6 - CH1(5)",
                       "EStop Level 7" := "E-STOP L7 - CH1(5)",
                       "EStop Level 8" := "E-STOP L8 - CH1(5)",
                       Bypass := "Bypass_Safe".Remote_Panel_5,
                       Overhang_Left := "Overhang_IO_DB".ECnv_5.Left,
                       Overhang_Right := "Overhang_IO_DB".ECnv_5.Right,
                       "STO VTD - CH1" => "STO VTD - CH1(5)",
                       "STO VTD - CH2" => "STO VTD - CH2(5)",
                       "STO CONVEYOR VTD - CH1" => "STO CONVEYOR VTD - CH1(5)",
                       "STO CONVEYOR VTD - CH2" => "STO CONVEYOR VTD - CH2(5)",
                       "STO CNV VFD (Level 1,2,3 - Side1) - CH1" => "STO CNV VFD (Level 1,2,3 - Side1) - CH1(5)",
                       "STO CNV VFD (Level 1,2,3 - Side1) - CH2" => "STO CNV VFD (Level 1,2,3 - Side1) - CH2(5)",
                       "STO CNV VFD (Level 4,5,6 - Side1) - CH1" => "STO CNV VFD (Level 4,5,6 - Side1) - CH1(5)",
                       "STO CNV VFD (Level 4,5,6 - Side1) - CH2" => "STO CNV VFD (Level 4,5,6 - Side1) - CH2(5)",
                       "STO CNV VFD (Level 7,8 - Side1) - CH1" => "STO CNV VFD (Level 7,8 - Side1) - CH1(5)",
                       "STO CNV VFD (Level 7,8 - Side1) - CH2" => "STO CNV VFD (Level 7,8 - Side1) - CH2(5)",
                       "Power Enable Safety Stopper Conveyors (Level 1,2,3 - Side1) - CH1" => "Power Enable Safety Stopper Conveyors (Level 1,2,3 - Side1) - CH1(5)",
                       "Power Enable Safety Stopper Conveyors (Level 1,2,3 - Side1) - CH2" => "Power Enable Safety Stopper Conveyors (Level 1,2,3 - Side1) - CH2(5)",
                       "Power Enable Safety Stopper Conveyors (Level 4,5,6 - Side1) - CH1" => "Power Enable Safety Stopper Conveyors (Level 4,5,6 - Side1) - CH1(5)",
                       "Power Enable Safety Stopper Conveyors (Level 4,5,6 - Side1) - CH2" => "Power Enable Safety Stopper Conveyors (Level 4,5,6 - Side1) - CH2(5)",
                       "Power Enable Safety Stopper Conveyors (Level 7,8 - Side1) - CH1" => "Power Enable Safety Stopper Conveyors (Level 7,8 - Side1) - CH1(5)",
                       "Power Enable Safety Stopper Conveyors (Level 7,8 - Side1) - CH2" => "Power Enable Safety Stopper Conveyors (Level 7,8 - Side1) - CH2(5)",
                       "VTU Hoist Brake Sfty Enable - CH1" => "VTU HOIST BRAKE SAFETY ENABLE 1(5)",
                       "VTU Hoist Brake Sfty Enable - CH2" => "VTU HOIST BRAKE SAFETY ENABLE 2(5)");
END_REGION

REGION Network 9: ESTOP LEVEL PANELS
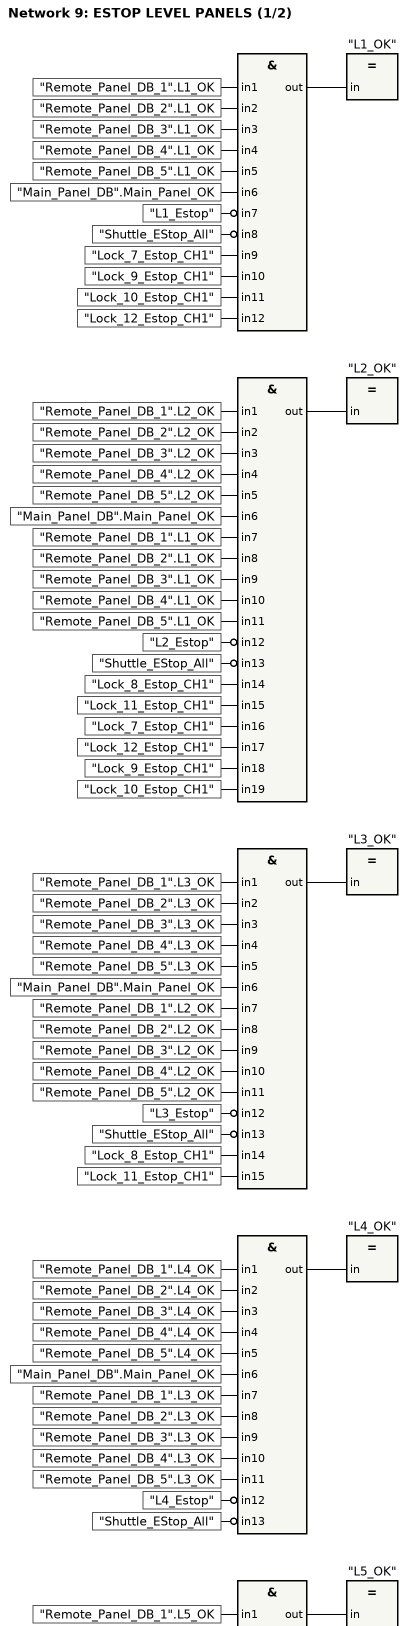
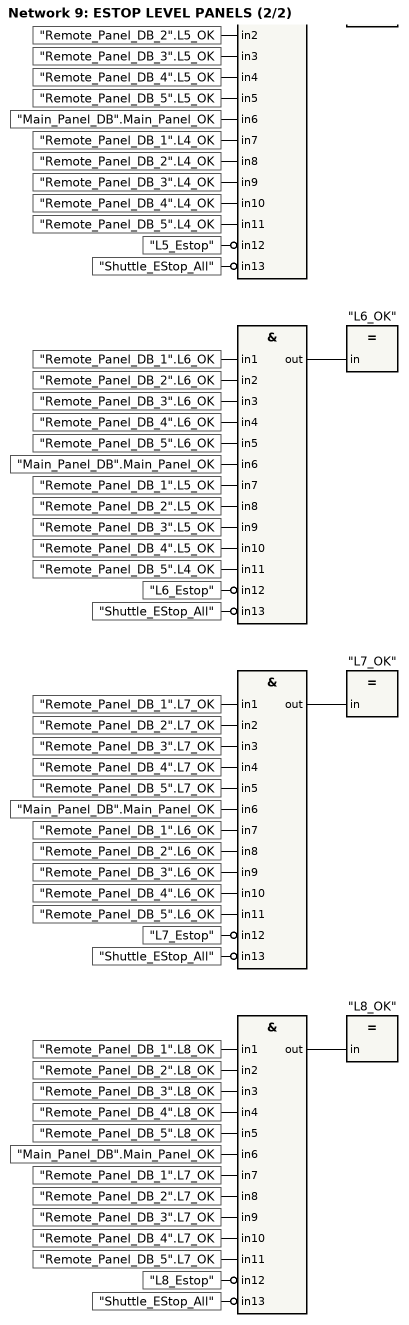
   "L1_OK" := "Remote_Panel_DB_1".L1_OK AND "Remote_Panel_DB_2".L1_OK AND "Remote_Panel_DB_3".L1_OK AND "Remote_Panel_DB_4".L1_OK AND "Remote_Panel_DB_5".L1_OK AND "Main_Panel_DB".Main_Panel_OK AND NOT "L1_Estop" AND NOT "Shuttle_EStop_All" AND "Lock_7_Estop_CH1" AND "Lock_9_Estop_CH1" AND "Lock_10_Estop_CH1" AND "Lock_12_Estop_CH1";
   "L2_OK" := "Remote_Panel_DB_1".L2_OK AND "Remote_Panel_DB_2".L2_OK AND "Remote_Panel_DB_3".L2_OK AND "Remote_Panel_DB_4".L2_OK AND "Remote_Panel_DB_5".L2_OK AND "Main_Panel_DB".Main_Panel_OK AND "Remote_Panel_DB_1".L1_OK AND "Remote_Panel_DB_2".L1_OK AND "Remote_Panel_DB_3".L1_OK AND "Remote_Panel_DB_4".L1_OK AND "Remote_Panel_DB_5".L1_OK AND NOT "L2_Estop" AND NOT "Shuttle_EStop_All" AND "Lock_8_Estop_CH1" AND "Lock_11_Estop_CH1" AND "Lock_7_Estop_CH1" AND "Lock_12_Estop_CH1" AND "Lock_9_Estop_CH1" AND "Lock_10_Estop_CH1";
   "L3_OK" := "Remote_Panel_DB_1".L3_OK AND "Remote_Panel_DB_2".L3_OK AND "Remote_Panel_DB_3".L3_OK AND "Remote_Panel_DB_4".L3_OK AND "Remote_Panel_DB_5".L3_OK AND "Main_Panel_DB".Main_Panel_OK AND "Remote_Panel_DB_1".L2_OK AND "Remote_Panel_DB_2".L2_OK AND "Remote_Panel_DB_3".L2_OK AND "Remote_Panel_DB_4".L2_OK AND "Remote_Panel_DB_5".L2_OK AND NOT "L3_Estop" AND NOT "Shuttle_EStop_All" AND "Lock_8_Estop_CH1" AND "Lock_11_Estop_CH1";
   "L4_OK" := "Remote_Panel_DB_1".L4_OK AND "Remote_Panel_DB_2".L4_OK AND "Remote_Panel_DB_3".L4_OK AND "Remote_Panel_DB_4".L4_OK AND "Remote_Panel_DB_5".L4_OK AND "Main_Panel_DB".Main_Panel_OK AND "Remote_Panel_DB_1".L3_OK AND "Remote_Panel_DB_2".L3_OK AND "Remote_Panel_DB_3".L3_OK AND "Remote_Panel_DB_4".L3_OK AND "Remote_Panel_DB_5".L3_OK AND NOT "L4_Estop" AND NOT "Shuttle_EStop_All";
   "L5_OK" := "Remote_Panel_DB_1".L5_OK AND "Remote_Panel_DB_2".L5_OK AND "Remote_Panel_DB_3".L5_OK AND "Remote_Panel_DB_4".L5_OK AND "Remote_Panel_DB_5".L5_OK AND "Main_Panel_DB".Main_Panel_OK AND "Remote_Panel_DB_1".L4_OK AND "Remote_Panel_DB_2".L4_OK AND "Remote_Panel_DB_3".L4_OK AND "Remote_Panel_DB_4".L4_OK AND "Remote_Panel_DB_5".L4_OK AND NOT "L5_Estop" AND NOT "Shuttle_EStop_All";
   "L6_OK" := "Remote_Panel_DB_1".L6_OK AND "Remote_Panel_DB_2".L6_OK AND "Remote_Panel_DB_3".L6_OK AND "Remote_Panel_DB_4".L6_OK AND "Remote_Panel_DB_5".L6_OK AND "Main_Panel_DB".Main_Panel_OK AND "Remote_Panel_DB_1".L5_OK AND "Remote_Panel_DB_2".L5_OK AND "Remote_Panel_DB_3".L5_OK AND "Remote_Panel_DB_4".L5_OK AND "Remote_Panel_DB_5".L4_OK AND NOT "L6_Estop" AND NOT "Shuttle_EStop_All";
   "L7_OK" := "Remote_Panel_DB_1".L7_OK AND "Remote_Panel_DB_2".L7_OK AND "Remote_Panel_DB_3".L7_OK AND "Remote_Panel_DB_4".L7_OK AND "Remote_Panel_DB_5".L7_OK AND "Main_Panel_DB".Main_Panel_OK AND "Remote_Panel_DB_1".L6_OK AND "Remote_Panel_DB_2".L6_OK AND "Remote_Panel_DB_3".L6_OK AND "Remote_Panel_DB_4".L6_OK AND "Remote_Panel_DB_5".L6_OK AND NOT "L7_Estop" AND NOT "Shuttle_EStop_All";
   "L8_OK" := "Remote_Panel_DB_1".L8_OK AND "Remote_Panel_DB_2".L8_OK AND "Remote_Panel_DB_3".L8_OK AND "Remote_Panel_DB_4".L8_OK AND "Remote_Panel_DB_5".L8_OK AND "Main_Panel_DB".Main_Panel_OK AND "Remote_Panel_DB_1".L7_OK AND "Remote_Panel_DB_2".L7_OK AND "Remote_Panel_DB_3".L7_OK AND "Remote_Panel_DB_4".L7_OK AND "Remote_Panel_DB_5".L7_OK AND NOT "L8_Estop" AND NOT "Shuttle_EStop_All";
END_REGION

REGION Network 10: LOCKS
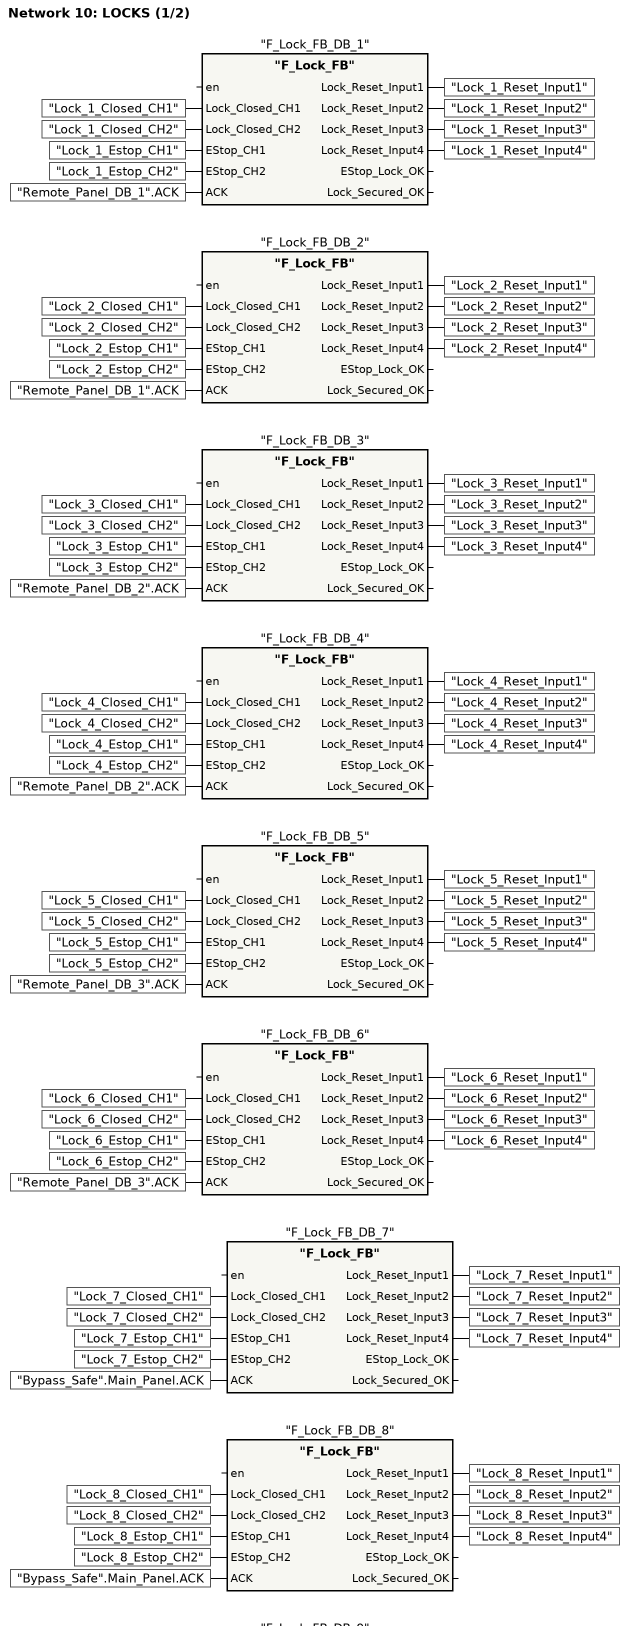
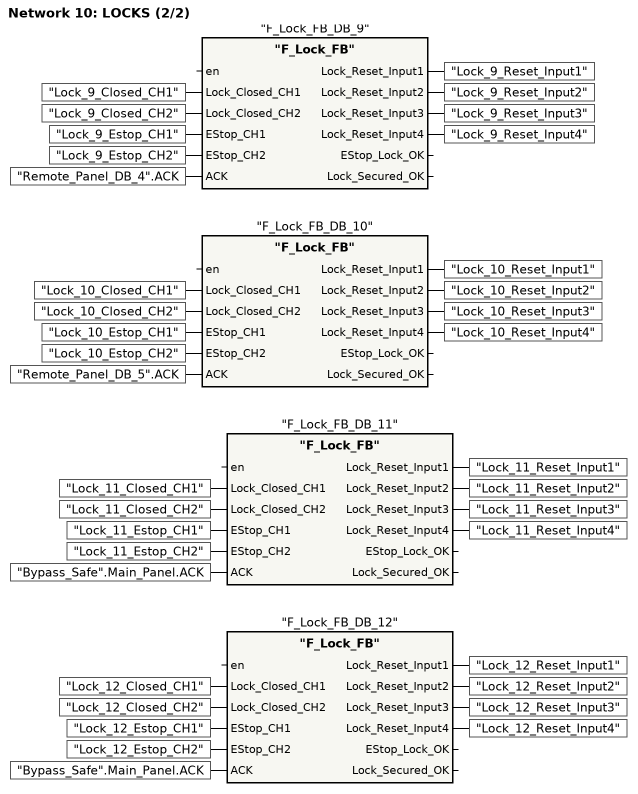
   "F_Lock_FB_DB_1"(Lock_Closed_CH1 := "Lock_1_Closed_CH1",   // "F_Lock_FB"
                    Lock_Closed_CH2 := "Lock_1_Closed_CH2",
                    EStop_CH1 := "Lock_1_Estop_CH1",
                    EStop_CH2 := "Lock_1_Estop_CH2",
                    ACK := "Remote_Panel_DB_1".ACK,
                    Lock_Reset_Input1 => "Lock_1_Reset_Input1",
                    Lock_Reset_Input2 => "Lock_1_Reset_Input2",
                    Lock_Reset_Input3 => "Lock_1_Reset_Input3",
                    Lock_Reset_Input4 => "Lock_1_Reset_Input4");
   "F_Lock_FB_DB_2"(Lock_Closed_CH1 := "Lock_2_Closed_CH1",   // "F_Lock_FB"
                    Lock_Closed_CH2 := "Lock_2_Closed_CH2",
                    EStop_CH1 := "Lock_2_Estop_CH1",
                    EStop_CH2 := "Lock_2_Estop_CH2",
                    ACK := "Remote_Panel_DB_1".ACK,
                    Lock_Reset_Input1 => "Lock_2_Reset_Input1",
                    Lock_Reset_Input2 => "Lock_2_Reset_Input2",
                    Lock_Reset_Input3 => "Lock_2_Reset_Input3",
                    Lock_Reset_Input4 => "Lock_2_Reset_Input4");
   "F_Lock_FB_DB_3"(Lock_Closed_CH1 := "Lock_3_Closed_CH1",   // "F_Lock_FB"
                    Lock_Closed_CH2 := "Lock_3_Closed_CH2",
                    EStop_CH1 := "Lock_3_Estop_CH1",
                    EStop_CH2 := "Lock_3_Estop_CH2",
                    ACK := "Remote_Panel_DB_2".ACK,
                    Lock_Reset_Input1 => "Lock_3_Reset_Input1",
                    Lock_Reset_Input2 => "Lock_3_Reset_Input2",
                    Lock_Reset_Input3 => "Lock_3_Reset_Input3",
                    Lock_Reset_Input4 => "Lock_3_Reset_Input4");
   "F_Lock_FB_DB_4"(Lock_Closed_CH1 := "Lock_4_Closed_CH1",   // "F_Lock_FB"
                    Lock_Closed_CH2 := "Lock_4_Closed_CH2",
                    EStop_CH1 := "Lock_4_Estop_CH1",
                    EStop_CH2 := "Lock_4_Estop_CH2",
                    ACK := "Remote_Panel_DB_2".ACK,
                    Lock_Reset_Input1 => "Lock_4_Reset_Input1",
                    Lock_Reset_Input2 => "Lock_4_Reset_Input2",
                    Lock_Reset_Input3 => "Lock_4_Reset_Input3",
                    Lock_Reset_Input4 => "Lock_4_Reset_Input4");
   "F_Lock_FB_DB_5"(Lock_Closed_CH1 := "Lock_5_Closed_CH1",   // "F_Lock_FB"
                    Lock_Closed_CH2 := "Lock_5_Closed_CH2",
                    EStop_CH1 := "Lock_5_Estop_CH1",
                    EStop_CH2 := "Lock_5_Estop_CH2",
                    ACK := "Remote_Panel_DB_3".ACK,
                    Lock_Reset_Input1 => "Lock_5_Reset_Input1",
                    Lock_Reset_Input2 => "Lock_5_Reset_Input2",
                    Lock_Reset_Input3 => "Lock_5_Reset_Input3",
                    Lock_Reset_Input4 => "Lock_5_Reset_Input4");
   "F_Lock_FB_DB_6"(Lock_Closed_CH1 := "Lock_6_Closed_CH1",   // "F_Lock_FB"
                    Lock_Closed_CH2 := "Lock_6_Closed_CH2",
                    EStop_CH1 := "Lock_6_Estop_CH1",
                    EStop_CH2 := "Lock_6_Estop_CH2",
                    ACK := "Remote_Panel_DB_3".ACK,
                    Lock_Reset_Input1 => "Lock_6_Reset_Input1",
                    Lock_Reset_Input2 => "Lock_6_Reset_Input2",
                    Lock_Reset_Input3 => "Lock_6_Reset_Input3",
                    Lock_Reset_Input4 => "Lock_6_Reset_Input4");
   "F_Lock_FB_DB_7"(Lock_Closed_CH1 := "Lock_7_Closed_CH1",   // "F_Lock_FB"
                    Lock_Closed_CH2 := "Lock_7_Closed_CH2",
                    EStop_CH1 := "Lock_7_Estop_CH1",
                    EStop_CH2 := "Lock_7_Estop_CH2",
                    ACK := "Bypass_Safe".Main_Panel.ACK,
                    Lock_Reset_Input1 => "Lock_7_Reset_Input1",
                    Lock_Reset_Input2 => "Lock_7_Reset_Input2",
                    Lock_Reset_Input3 => "Lock_7_Reset_Input3",
                    Lock_Reset_Input4 => "Lock_7_Reset_Input4");
   "F_Lock_FB_DB_8"(Lock_Closed_CH1 := "Lock_8_Closed_CH1",   // "F_Lock_FB"
                    Lock_Closed_CH2 := "Lock_8_Closed_CH2",
                    EStop_CH1 := "Lock_8_Estop_CH1",
                    EStop_CH2 := "Lock_8_Estop_CH2",
                    ACK := "Bypass_Safe".Main_Panel.ACK,
                    Lock_Reset_Input1 => "Lock_8_Reset_Input1",
                    Lock_Reset_Input2 => "Lock_8_Reset_Input2",
                    Lock_Reset_Input3 => "Lock_8_Reset_Input3",
                    Lock_Reset_Input4 => "Lock_8_Reset_Input4");
   "F_Lock_FB_DB_9"(Lock_Closed_CH1 := "Lock_9_Closed_CH1",   // "F_Lock_FB"
                    Lock_Closed_CH2 := "Lock_9_Closed_CH2",
                    EStop_CH1 := "Lock_9_Estop_CH1",
                    EStop_CH2 := "Lock_9_Estop_CH2",
                    ACK := "Remote_Panel_DB_4".ACK,
                    Lock_Reset_Input1 => "Lock_9_Reset_Input1",
                    Lock_Reset_Input2 => "Lock_9_Reset_Input2",
                    Lock_Reset_Input3 => "Lock_9_Reset_Input3",
                    Lock_Reset_Input4 => "Lock_9_Reset_Input4");
   "F_Lock_FB_DB_10"(Lock_Closed_CH1 := "Lock_10_Closed_CH1",   // "F_Lock_FB"
                     Lock_Closed_CH2 := "Lock_10_Closed_CH2",
                     EStop_CH1 := "Lock_10_Estop_CH1",
                     EStop_CH2 := "Lock_10_Estop_CH2",
                     ACK := "Remote_Panel_DB_5".ACK,
                     Lock_Reset_Input1 => "Lock_10_Reset_Input1",
                     Lock_Reset_Input2 => "Lock_10_Reset_Input2",
                     Lock_Reset_Input3 => "Lock_10_Reset_Input3",
                     Lock_Reset_Input4 => "Lock_10_Reset_Input4");
   "F_Lock_FB_DB_11"(Lock_Closed_CH1 := "Lock_11_Closed_CH1",   // "F_Lock_FB"
                     Lock_Closed_CH2 := "Lock_11_Closed_CH2",
                     EStop_CH1 := "Lock_11_Estop_CH1",
                     EStop_CH2 := "Lock_11_Estop_CH2",
                     ACK := "Bypass_Safe".Main_Panel.ACK,
                     Lock_Reset_Input1 => "Lock_11_Reset_Input1",
                     Lock_Reset_Input2 => "Lock_11_Reset_Input2",
                     Lock_Reset_Input3 => "Lock_11_Reset_Input3",
                     Lock_Reset_Input4 => "Lock_11_Reset_Input4");
   "F_Lock_FB_DB_12"(Lock_Closed_CH1 := "Lock_12_Closed_CH1",   // "F_Lock_FB"
                     Lock_Closed_CH2 := "Lock_12_Closed_CH2",
                     EStop_CH1 := "Lock_12_Estop_CH1",
                     EStop_CH2 := "Lock_12_Estop_CH2",
                     ACK := "Bypass_Safe".Main_Panel.ACK,
                     Lock_Reset_Input1 => "Lock_12_Reset_Input1",
                     Lock_Reset_Input2 => "Lock_12_Reset_Input2",
                     Lock_Reset_Input3 => "Lock_12_Reset_Input3",
                     Lock_Reset_Input4 => "Lock_12_Reset_Input4");
END_REGION

REGION Network 11: Safety OK
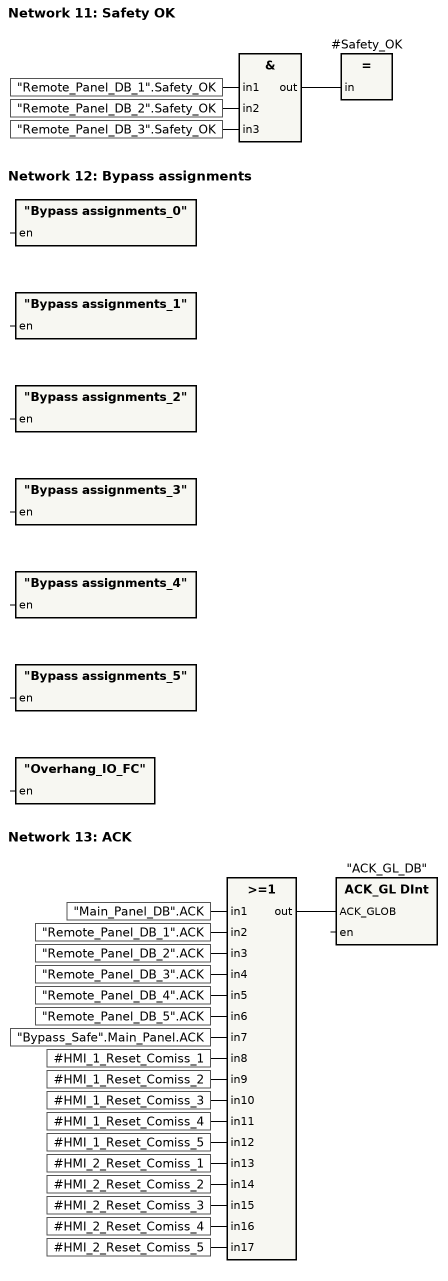
   #Safety_OK := "Remote_Panel_DB_1".Safety_OK AND "Remote_Panel_DB_2".Safety_OK AND "Remote_Panel_DB_3".Safety_OK;
END_REGION

REGION Network 12: Bypass assignments
   "Bypass assignments_0"();
   "Bypass assignments_1"();
   "Bypass assignments_2"();
   "Bypass assignments_3"();
   "Bypass assignments_4"();
   "Bypass assignments_5"();
   "Overhang_IO_FC"();
END_REGION

REGION Network 13: ACK
   "ACK_GL_DB"(ACK_GLOB := "Main_Panel_DB".ACK OR "Remote_Panel_DB_1".ACK OR "Remote_Panel_DB_2".ACK OR "Remote_Panel_DB_3".ACK OR "Remote_Panel_DB_4".ACK OR "Remote_Panel_DB_5".ACK OR "Bypass_Safe".Main_Panel.ACK OR #HMI_1_Reset_Comiss_1 OR #HMI_1_Reset_Comiss_2 OR #HMI_1_Reset_Comiss_3 OR #HMI_1_Reset_Comiss_4 OR #HMI_1_Reset_Comiss_5 OR #HMI_2_Reset_Comiss_1 OR #HMI_2_Reset_Comiss_2 OR #HMI_2_Reset_Comiss_3 OR #HMI_2_Reset_Comiss_4 OR #HMI_2_Reset_Comiss_5);   // ACK_GL
END_REGION

REGION Network 14: RESET PLC HMI
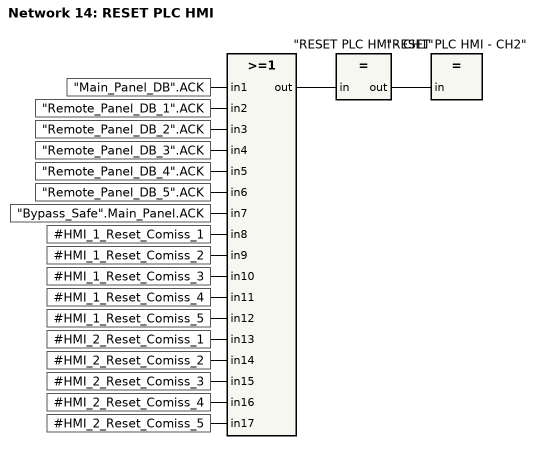
   "RESET PLC HMI - CH1" := "Main_Panel_DB".ACK OR "Remote_Panel_DB_1".ACK OR "Remote_Panel_DB_2".ACK OR "Remote_Panel_DB_3".ACK OR "Remote_Panel_DB_4".ACK OR "Remote_Panel_DB_5".ACK OR "Bypass_Safe".Main_Panel.ACK OR #HMI_1_Reset_Comiss_1 OR #HMI_1_Reset_Comiss_2 OR #HMI_1_Reset_Comiss_3 OR #HMI_1_Reset_Comiss_4 OR #HMI_1_Reset_Comiss_5 OR #HMI_2_Reset_Comiss_1 OR #HMI_2_Reset_Comiss_2 OR #HMI_2_Reset_Comiss_3 OR #HMI_2_Reset_Comiss_4 OR #HMI_2_Reset_Comiss_5;
   "RESET PLC HMI - CH2" := "RESET PLC HMI - CH1";
END_REGION
END_FUNCTION_BLOCK
